(* IEC 61131-3 sources: Codesys_IAP/Demo/PLC1/Magazijn Overzetter Simulatie Structured Text 2V1 - Leeg_tekst/Programma Structured Text/OverzetterClass, 7 files *)

(* ---- cycle.st ---- *)
(*#### DECLARATIE ####*)
// Datum : 17 december 2020, Auteur: Gerard Harkema
METHOD cycle
VAR
END_VAR
(*#### IMPLEMENTATIE ####*)
CASE eState OF

//	overzetterStates.idle :
	overzetterStates.ga_naar_links:
		IF IO.Ix_OverzetterIsLinks THEN
			IO.Qx_OverzetterLinks 		:= FALSE;
			IO.Qx_VacuumAan 			:= TRUE;
			eState 					:= overzetterStates.is_links;
		END_IF;
	overzetterStates.is_links:
		IF IO.Ix_VacuumAanwezig THEN
			IO.Qx_OverzetterRechts 	:= TRUE;
			eState					:= overzetterStates.ga_naar_rechts;
	END_IF
//	overzetterStates.vaccuum_aanzetten:
	overzetterStates.ga_naar_rechts:
		IF IO.Ix_OverzetterIsRechts THEN
			IO.Qx_OverzetterRechts := FALSE;
			IO.Qx_VacuumAan 		:= FALSE;
			IO.Qx_BekerLossen 		:= TRUE;
			eState := overzetterStates.is_rechts;
		END_IF
	overzetterStates.is_rechts:
		IF NOT IO.Ix_VacuumAanwezig THEN
			IO.Qx_BekerLossen 		:= FALSE;
			IO.Qx_OverzetterLinks 	:= TRUE;
			eState 				:= overzetterStates.ga_naar_midden;
		END_IF
//	overzetterStates.vaccuum_lossen:
	overzetterStates.ga_naar_midden:
		IF timer.Q THEN
			IO.Qx_OverzetterLinks	:= FALSE;
			eState 				:= overzetterStates.is_midden;
			xKlaar 					:= TRUE;
		END_IF

	//overzetterStates.is_midden:
//	overzetterStates.error:
END_CASE

timer(IN:=(estate =overzetterStates.ga_naar_midden), PT:=T#2S);

(* ---- initialize.st ---- *)
(*#### DECLARATIE ####*)
// Datum : 17 december 2020, Auteur: Gerard Harkema
METHOD initialize
VAR_INPUT
	IORef		: REFERENCE TO overzetterIO;
END_VAR
(*#### IMPLEMENTATIE ####*)
IO							REF= IORef;

IO.Qx_BekerLossen			:= FALSE;
IO.Qx_VacuumAan				:= FALSE;
IO.Qx_OverzetterLinks		:= FALSE;
IO.Qx_OverzetterRechts		:= TRUE;
eState 						:= overzetterStates.ga_naar_rechts;

(* ---- isError.st ---- *)
(*#### DECLARATIE ####*)
// Datum : 17 december 2020, Auteur: Gerard Harkema
METHOD isError : BOOL
VAR_INPUT
END_VAR
(*#### IMPLEMENTATIE ####*)
isError := (eState = overzetterStates.error);

(* ---- isKlaar.st ---- *)
(*#### DECLARATIE ####*)
// Datum : 17 december 2020, Auteur: Gerard Harkema
METHOD isKlaar : BOOL
VAR_INPUT
END_VAR
(*#### IMPLEMENTATIE ####*)
isKlaar := xKlaar;

(* ---- noodstop.st ---- *)
(*#### DECLARATIE ####*)
// Datum : 17 december 2020, Auteur: Gerard Harkema
METHOD noodstop
VAR_INPUT
END_VAR
(*#### IMPLEMENTATIE ####*)
//Beker oppakken
IO.Qx_VacuumAan 			:=FALSE;
//Beker loslaten
IO.Qx_BekerLossen 			:=FALSE;
//Overzetter naar bekermagazijn
IO.Qx_OverzetterLinks 		:=FALSE;
//Overzetter naar sorteerpositie
IO.Qx_OverzetterRechts 	:=FALSE;

eState 				:= overzetterStates.error;

(* ---- reset.st ---- *)
(*#### DECLARATIE ####*)
// Datum : 17 december 2020, Auteur: Gerard Harkema
METHOD reset
VAR_INPUT
END_VAR
(*#### IMPLEMENTATIE ####*)
IO.Qx_BekerLossen			:= FALSE;
IO.Qx_VacuumAan				:= FALSE;
IO.Qx_OverzetterLinks		:= FALSE;
IO.Qx_OverzetterRechts		:= TRUE;
eState 						:= overzetterStates.ga_naar_rechts;
// Pas weer klaar als de ruststand bereikt is
xKlaar						:= FALSE;

(* ---- start.st ---- *)
(*#### DECLARATIE ####*)
// Datum : 17 december 2020, Auteur: Gerard Harkema
METHOD start : BOOL
VAR_INPUT
END_VAR
(*#### IMPLEMENTATIE ####*)
IF NOT (eState = overzetterStates.is_midden) THEN
	eState 				:= overzetterStates.error;
//	IO.Qx_BekerUitstoten 	:= FALSE;
	start 	:= TRUE; // Failed
	RETURN;
END_IF

xKlaar 					:= FALSE;
IO.Qx_OverzetterLinks 		:= TRUE;
eState 					:= overzetterStates.ga_naar_links;

start			:= FALSE; // oké
